(* Munsch command *)
TYPE ET_MUNSCH_CMD :
(
	ET_MUNSCH_CMD_NOCMD := 0,
	ET_MUNSCH_CMD_STARTHEAT := 1,
	ET_MUNSCH_CMD_STOPHEAT := 2,
	ET_MUNSCH_CMD_REQHEATSTATUS := 3,
	ET_MUNSCH_CMD_STARTEXTRUDER := 5,
	ET_MUNSCH_CMD_STOPEXTRUDER := 6,
	ET_MUNSCH_CMD_REQEXTRUDERSTATUS := 7,
	ET_MUNSCH_CMD_SETMATERIALTEMP := 9,
	ET_MUNSCH_CMD_REQMATERIALREFTEMP := 10,
	ET_MUNSCH_CMD_REQMATERIALACTTEMP := 11,
	ET_MUNSCH_CMD_SETAIRTEMP := 13,
	ET_MUNSCH_CMD_REQAIRREFTEMP := 14,
	ET_MUNSCH_CMD_REQAIRACTTEMP := 15,
	ET_MUNSCH_CMD_REQSTATUS := 20

);
END_TYPE

(* stored: Version 1.1.0.1, ProductVersion 3.1.4024.15
   DUT ET_MUNSCH_CMD: Id {829c7538-b7e6-4f60-945e-74c0e0b3ce20} *)
